Fanuc KAREL source: KA00159.KL

PROGRAM KA00159
%NOLOCKGROUP
VAR
  SRC: ARRAY[4] OF REAL
  DST: ARRAY[4] OF SHORT
BEGIN
  DST = SRC
END KA00159
